// TIA Portal V20 export
Screen "Call_ServiceButtons_1"  1276x673
  ScreenItem "Title_OPMode1_ScreenOverview_X390_Y2" at 5,7 size 1262x30  Type=HmiTextBox
  ScreenItem "Faceplate container_5" at 0,33 size 622x206  Type=HmiFaceplateContainer
  ScreenItem "Text box_5" at 0,0 size 622x30  Type=HmiTextBox
  ScreenItem "Faceplate container_7" at 0,33 size 622x206  Type=HmiFaceplateContainer
  ScreenItem "Text box_7" at 0,0 size 622x30  Type=HmiTextBox
  ScreenItem "Faceplate container_8" at 0,33 size 622x206  Type=HmiFaceplateContainer
  ScreenItem "Text box_8" at 0,0 size 622x30  Type=HmiTextBox
  ScreenItem "Faceplate container_3" at 646,286 size 619x179  Type=HmiFaceplateContainer
  ScreenItem "Text box_3" at 645,255 size 622x30  Type=HmiTextBox
  ScreenItem "Faceplate container_4" at 646,496 size 619x179  Type=HmiFaceplateContainer
  ScreenItem "Text box_4" at 645,466 size 622x30  Type=HmiTextBox
  ScreenItem "Faceplate container_6" at 14,74 size 619x179  Type=HmiFaceplateContainer
  ScreenItem "Text box_6" at 13,41 size 622x30  Type=HmiTextBox
  ScreenItem "Faceplate container_9" at 646,74 size 619x179  Type=HmiFaceplateContainer
  ScreenItem "Text box_9" at 648,41 size 622x30  Type=HmiTextBox
  ScreenItem "Faceplate container_1" at 14,285 size 619x179  Type=HmiFaceplateContainer
  ScreenItem "Text box_1" at 13,254 size 622x30  Type=HmiTextBox
  ScreenItem "Faceplate container_2" at 14,496 size 619x179  Type=HmiFaceplateContainer
  ScreenItem "Text box_2" at 13,466 size 622x30  Type=HmiTextBox
  ScreenItem "Button_15" at 1170,8 size 98x31  Type=HmiButton
